(* PLC project TBEN_L5_PLC11.project, CODESYS CODESYS V3.5 SP21 Patch 1 *)
(* stored: creationDateTime 2026-11-07T15:22:03.2751678, modificationDateTime 2026-11-07T15:09:07.4034196 *)

(* global variable list GVL_IO *)
// Ngõ vào/ra DXP của TBEN-L5-PLC-11 (map trong Local_IO > DXP > I/O Mapping)
// Đầu nối: C4 = Ch8/Ch9, C5 = Ch10/Ch11, C6 = Ch12/Ch13, C7 = Ch14/Ch15
VAR_GLOBAL
    xQ_Ch8  : BOOL;   // ngõ ra DXP Ch8  (C4)
    xQ_Ch9  : BOOL;   // ngõ ra DXP Ch9  (C4)
    xQ_Ch10 : BOOL;   // ngõ ra DXP Ch10 (C5)
    xQ_Ch11 : BOOL;   // ngõ ra DXP Ch11 (C5)
    xQ_Ch12 : BOOL;   // ngõ ra DXP Ch12 (C6)
    xQ_Ch13 : BOOL;   // ngõ ra DXP Ch13 (C6)
    xQ_Ch14 : BOOL;   // ngõ ra DXP Ch14 (C7)
    xQ_Ch15 : BOOL;   // ngõ ra DXP Ch15 (C7)

    xI_Ch8  : BOOL;   // đọc lại mức tín hiệu DXP Ch8
    xI_Ch9  : BOOL;   // đọc lại mức tín hiệu DXP Ch9
    xI_Ch10 : BOOL;   // đọc lại mức tín hiệu DXP Ch10
    xI_Ch11 : BOOL;   // đọc lại mức tín hiệu DXP Ch11
    xI_Ch12 : BOOL;   // đọc lại mức tín hiệu DXP Ch12
    xI_Ch13 : BOOL;   // đọc lại mức tín hiệu DXP Ch13
    xI_Ch14 : BOOL;   // đọc lại mức tín hiệu DXP Ch14
    xI_Ch15 : BOOL;   // đọc lại mức tín hiệu DXP Ch15
END_VAR
